// TIA Portal V20 export
Screen "190FX2RhSliderFixtureLayout"  1276x673
  ScreenItem "Line_Header_X0_Y64" at 0,64 size 1276x0  Type=HmiLine
  ScreenItem "permanentareaborderrectangle" at 0,0 size 0x0  Type=HmiRectangle
  ScreenItem "Button_Back" at 2,2 size 90x60  Type=HmiButton
  ScreenItem "Move_Legend" at 1182,2 size 90x60  Type=HmiButton
  ScreenItem "Fusszeile_Button_ManualOPMode1_2" at 279,2 size 90x60  Type=HmiButton
  ScreenItem "文本域_3" at 1107,71 size 139x22  Type=HmiTextBox
  ScreenItem "文本域_1" at 1107,160 size 156x23  Type=HmiTextBox
  ScreenItem "文本域_2" at 1098,246 size 165x23  Type=HmiTextBox
  ScreenItem "文本域_22" at 1124,475 size 104x23  Type=HmiTextBox
  ScreenItem "Fusszeile_Button_ManualOPMode1_1" at 95,2 size 90x60  Type=HmiButton
  ScreenItem "Button_Back_1" at 1180,606 size 90x60  Type=HmiButton
  ScreenItem "Fusszeile_Button_ManualOPMode1_3" at 187,2 size 90x60  Type=HmiButton
  ScreenItem "Fusszeile_Button_ManualOPMode1_4" at 997,2 size 90x60  Type=HmiButton
  ScreenItem "Fusszeile_Button_ManualOPMode1_5" at 902,1 size 90x60  Type=HmiButton
  ScreenItem "文本域_14" at 936,-172 size 140x40  Type=HmiTextBox
  ScreenItem "Title_ScreenOverview_X390_Y2_1" at 384,5 size 510x57  Type=HmiTextBox
  ScreenItem "Graphic view_1" at 260,212 size 560x296  Type=HmiGraphicView
  ScreenItem "文本域_5" at -1,82 size 120x40  Type=HmiTextBox
  ScreenItem "文本域_27" at -1,126 size 120x40  Type=HmiTextBox
  ScreenItem "LSicar_Valve8Pos_LeftHomeRightWork_WithPB_5" at 1099,95 size 160x53  Type=HmiFaceplateContainer
  ScreenItem "LSicar_Valve8Pos_LeftHomeRightWork_WithPB_1" at 1099,183 size 160x53  Type=HmiFaceplateContainer
  ScreenItem "面板容器_22" at 1061,508 size 96x32  Type=HmiFaceplateContainer
  ScreenItem "面板容器_23" at 1171,508 size 96x32  Type=HmiFaceplateContainer
  ScreenItem "LSicar_Valve8Pos_LeftHomeRightWork_WithPB_2" at 1099,271 size 160x53  Type=HmiFaceplateContainer
  ScreenItem "文本域_21" at 350,99 size 140x40  Type=HmiTextBox
  ScreenItem "Line_4" at 234,225 size 239x36  Type=HmiLine
  ScreenItem "文本域_12" at 133,196 size 100x40  Type=HmiTextBox
  ScreenItem "Line_1" at 443,194 size 116x84  Type=HmiLine
  ScreenItem "文本域_6" at 873,196 size 140x40  Type=HmiTextBox
  ScreenItem "面板容器_1" at 875,237 size 144x51  Type=HmiFaceplateContainer
  ScreenItem "Line_2" at 672,209 size 193x80  Type=HmiLine
  ScreenItem "文本域_7" at 783,98 size 100x40  Type=HmiTextBox
  ScreenItem "Faceplate container_1" at 803,139 size 59x45  Type=HmiFaceplateContainer
  ScreenItem "Line_3" at 663,156 size 138x105  Type=HmiLine
  ScreenItem "文本域_8" at 844,392 size 100x40  Type=HmiTextBox
  ScreenItem "Faceplate container_2" at 864,433 size 59x45  Type=HmiFaceplateContainer
  ScreenItem "Line_5" at 645,300 size 194x108  Type=HmiLine
  ScreenItem "文本域_9" at 594,522 size 100x40  Type=HmiTextBox
  ScreenItem "Faceplate container_3" at 614,562 size 59x45  Type=HmiFaceplateContainer
  ScreenItem "Line_6" at 592,338 size 50x180  Type=HmiLine
  ScreenItem "文本域_10" at 133,392 size 100x40  Type=HmiTextBox
  ScreenItem "Faceplate container_4" at 153,433 size 59x45  Type=HmiFaceplateContainer
  ScreenItem "Line_7" at 233,302 size 252x98  Type=HmiLine
  ScreenItem "文本域_13" at 540,99 size 140x40  Type=HmiTextBox
  ScreenItem "Line_9" at 594,187 size 9x110  Type=HmiLine
  ScreenItem "文本域_15" at 373,522 size 100x40  Type=HmiTextBox
  ScreenItem "Faceplate container_5" at 393,562 size 59x45  Type=HmiFaceplateContainer
  ScreenItem "Line_10" at 439,342 size 89x176  Type=HmiLine
  ScreenItem "Faceplate container_6" at 153,237 size 59x45  Type=HmiFaceplateContainer
  ScreenItem "面板容器_8" at 352,143 size 144x51  Type=HmiFaceplateContainer
  ScreenItem "面板容器_4" at 543,143 size 144x51  Type=HmiFaceplateContainer
  ScreenItem "面板容器_2" at 1090,4 size 88x58  Type=HmiFaceplateContainer
  ScreenItem "OPMode1_Blocked" at 1164,6 size 14x14  Type=HmiGraphicView
  ScreenItem "OPMode4_Foreground_Blocked" at 1089,2 size 88x58  Type=HmiGraphicView
